// TIA Portal V21 export
TYPE "Motor"
// A motor, assigned to a ProDiag function block where it is used.
   STRUCT
      running : Bool;
      tripped : Bool;
      ready : Bool;
      speed : Int;
   END_STRUCT;
END_TYPE
